// TIA Portal V19 export
TYPE "EM04_Input"
   STRUCT
      Cmds { S7_SetPoint := 'True'} : "EM_Input";
      CtrlMode : Int;   // 0=Off, 1=Inyeccion por tiempo, 2=Carga por nivel
      SelectedValveIndex : Int;   // Valvula de insumo seleccionada (1..NUM_VLV)
      InjectionTime : Time := T#3S;
      TargetLevelSP : Real;
      LevelFilter : Time := T#3S;
      LevelTimeout : Time := T#20M;
      LevelValid : Bool := TRUE;
      LevelInterlock : Bool;
   END_STRUCT;
END_TYPE
